Yaskawa INFORM job: DEMO_BUTTON_REPEAT.JBI

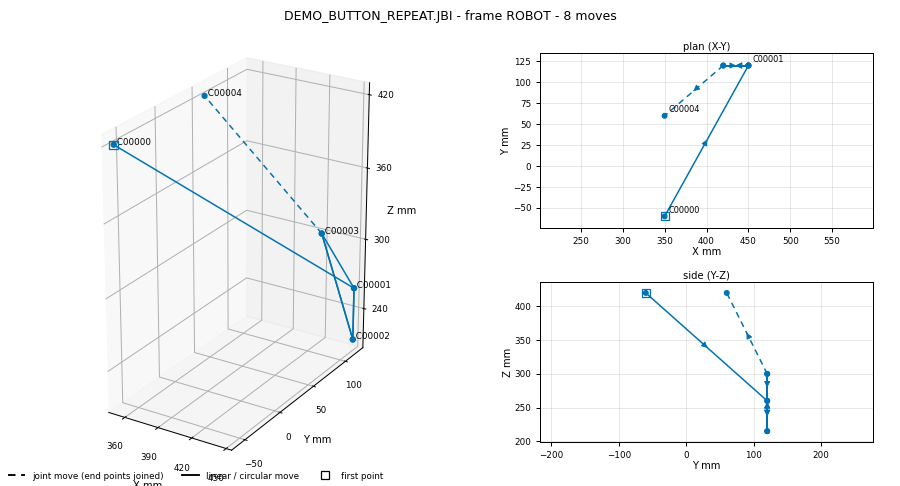
[picture p0: tool path of DEMO_BUTTON_REPEAT.JBI in frame ROBOT, 8 of 8 moves have a stored position in this frame; points joined in program order, loops and branches not executed]
/JOB
//NAME DEMO_BUTTON_REPEAT
//POS
///NPOS 5,0,0,0,0,0
///TOOL 0
///POSTYPE ROBOT
///RECTAN
///RCONF 0,0,0,0,0,0,0,0
C00000=350.000,-60.000,420.000,180.00,0.00,0.00
C00001=450.000,120.000,260.000,180.00,0.00,0.00
C00002=450.000,120.000,215.000,180.00,0.00,0.00
C00003=420.000,120.000,300.000,180.00,0.00,0.00
C00004=350.000,60.000,420.000,180.00,0.00,0.00
//INST
///DATE 2026/11/03 20:00
///ATTR SC,RW
///GROUP1 RB1
NOP
'SYNTHETIC DEMO JOB - NOT A REAL ROBOT JOB
MOVJ C00000 VJ=25.00
MOVL C00001 V=150.0
MOVL C00002 V=30.0
MOVL C00003 V=150.0
MOVL C00001 V=150.0
MOVL C00002 V=30.0
MOVL C00003 V=150.0
MOVJ C00004 VJ=25.00
END
